// TIA Portal V21 export
DATA_BLOCK "IDB_AnaDoubleCall"   // DB9
// stored: InstanceOfName FB_AnaDoubleCall, InstanceOfType FB
"FB_AnaDoubleCall"
   // VAR_INPUT
   //    PulseA : Bool;
   //    PulseB : Bool;
   // END_VAR
   // VAR_OUTPUT
   //    Count : Int;
   // END_VAR
   // VAR
   //    PartCounter { S7_SetPoint := 'True'} : CTU_INT;
   // END_VAR
BEGIN
END_DATA_BLOCK
